(* IEC 61131-3 sources: avi-aoi-management/scripts/ai-eval/ngau-nhien/kho/st-tv3-nhap-nhay/khung/src, 1 file *)

(* ---- NhapNhay.st ---- *)
FUNCTION_BLOCK NhapNhay
VAR_INPUT
    BAT : BOOL;
    T_SANG : TIME;
    T_TOI : TIME;
END_VAR
VAR_OUTPUT
    DEN : BOOL;
END_VAR
    (* TODO: cài đặt theo đề bài, dùng TON *)
    DEN := BAT;
END_FUNCTION_BLOCK
